Universal Robots PolyScope program: program_3.urp

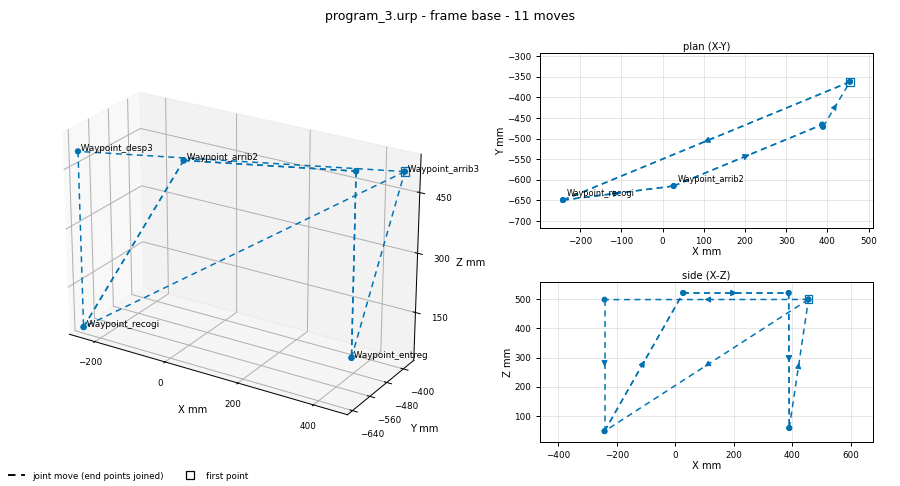
[picture p0: tool path of program_3.urp in frame base, 11 of 11 moves have a stored position in this frame; points joined in program order, loops and branches not executed]
Program program_3 (installation=default directory=/ursim/programs createdIn=3.15.8.106339 lastSavedIn=3.15.8.106339 robotSerialNumber=2018359999)
Calibrated DH parameters: a=[0, -0.425, -0.39225, 0, 0, 0]; d=[0.089159, 0, 0, 0.10915, 0.09465, 0.0823]; alpha=[1.570796, 0, 0, 1.570796, -1.570796, 0]; deltaTheta=[0, 0, 0, 0, 0, 0]
Robot Program (runOnlyOnce=false)
  MoveJ speed 60 deg/s, acceleration 80 deg/s^2 (useActiveTCP=true)
    Waypoint Waypoint_arrib3: TCP in base x=454.738 y=-362.048 z=498.534 mm, rx=-0.0012 ry=3.1165 rz=0.0387 rad; joints [-27.98, -102.369, -66.532, -100.508, 91.926, 61.985] deg
    Waypoint Waypoint_recogi: TCP in base x=-242.045 y=-649.292 z=48.33 mm, rx=-0.0012 ry=3.1165 rz=0.0387 rad; joints [-101.516, -134.482, -86.847, -50.351, 91.112, -11.577] deg
  Set DigitalOutput pin=digital_out[0]; digitalValue=1
  MoveJ speed 60 deg/s, acceleration 80 deg/s^2 (useActiveTCP=true)
    Waypoint Waypoint_arrib2: TCP in base x=26.637 y=-615.024 z=520.757 mm, rx=-0.0012 ry=3.1163 rz=0.0389 rad; joints [-77.539, -108.915, -54.252, -107.92, 91.71, 12.4] deg
    Waypoint Waypoint_despla: TCP in base x=387.077 y=-466.089 z=520.757 mm, rx=-0.0012 ry=3.1163 rz=0.0389 rad; joints [-40.191, -106.997, -57.155, -105.675, 92.019, 49.767] deg
    Waypoint Waypoint_entreg: TCP in base x=389.216 y=-471.264 z=59.159 mm, rx=-0.0012 ry=3.1163 rz=0.0389 rad; joints [-40.436, -125.554, -102.95, -41.332, 92.019, 49.522] deg
  Set DigitalOutput pin=digital_out[0]; digitalValue=0
  Set DigitalOutput pin=digital_out[0]; digitalValue=1
  MoveJ speed 60 deg/s, acceleration 80 deg/s^2 (useActiveTCP=true)
    Waypoint Waypoint_arrib3: TCP in base x=454.738 y=-362.048 z=498.534 mm, rx=-0.0012 ry=3.1165 rz=0.0387 rad; joints [-27.98, -102.369, -66.532, -100.508, 91.926, 61.985] deg
    Waypoint Waypoint_desp3: TCP in base x=-242.045 y=-649.292 z=497.929 mm, rx=-0.0012 ry=3.1165 rz=0.0387 rad; joints [-101.516, -121.643, -38.696, -111.341, 91.112, -11.577] deg
    Waypoint Waypoint_recogi: TCP in base x=-242.045 y=-649.292 z=48.33 mm, rx=-0.0012 ry=3.1165 rz=0.0387 rad; joints [-101.516, -134.482, -86.847, -50.351, 91.112, -11.577] deg
  Set DigitalOutput pin=digital_out[0]; digitalValue=0
  Set DigitalOutput pin=digital_out[0]; digitalValue=1
  MoveJ speed 60 deg/s, acceleration 80 deg/s^2 (useActiveTCP=true)
    Waypoint Waypoint_arrib2: TCP in base x=26.637 y=-615.024 z=520.757 mm, rx=-0.0012 ry=3.1163 rz=0.0389 rad; joints [-77.539, -108.915, -54.252, -107.92, 91.71, 12.4] deg
    Waypoint Waypoint_despla: TCP in base x=387.077 y=-466.089 z=520.757 mm, rx=-0.0012 ry=3.1163 rz=0.0389 rad; joints [-40.191, -106.997, -57.155, -105.675, 92.019, 49.767] deg
    Waypoint Waypoint_entreg: TCP in base x=389.216 y=-471.264 z=59.159 mm, rx=-0.0012 ry=3.1163 rz=0.0389 rad; joints [-40.436, -125.554, -102.95, -41.332, 92.019, 49.522] deg
  Set DigitalOutput pin=digital_out[0]; digitalValue=0
